// TIA Portal V19 export
DATA_BLOCK "ALL_PUMPS_DB"   // DB13
// stored: InstanceOfName ALL_PUMPS, InstanceOfType FB
"ALL_PUMPS"
   // VAR
   //    PUMP_FB1_CP01 { S7_SetPoint := 'True'} : "PUMP_FB1";
   //    PUMP_FB1_AG01 { S7_SetPoint := 'True'} : "PUMP_FB1";
   //    PUMP_FB1_CHS_CP01 { S7_SetPoint := 'True'} : "PUMP_FB1";
   //    PUMP_FB1_CHS_CP02 { S7_SetPoint := 'True'} : "PUMP_FB1";
   //    PUMP_FB1_CHS_CP03 { S7_SetPoint := 'True'} : "PUMP_FB1";
   //    PUMP_FB1_R2_CP01 { S7_SetPoint := 'True'} : "PUMP_FB1";
   //    PUMP_FB1_R2_AG01 { S7_SetPoint := 'True'} : "PUMP_FB1";
   //    PUMP_FB1_R3_CP01 { S7_SetPoint := 'True'} : "PUMP_FB1";
   //    PUMP_FB1_R3_AG01 { S7_SetPoint := 'True'} : "PUMP_FB1";
   //    PUMP_FB1_R4_CP01 { S7_SetPoint := 'True'} : "PUMP_FB1";
   //    PUMP_FB1_R4_AG01 { S7_SetPoint := 'True'} : "PUMP_FB1";
   //    PUMP_FB1_R5_CP01 { S7_SetPoint := 'True'} : "PUMP_FB1";
   //    PUMP_FB1_R5_AG01 { S7_SetPoint := 'True'} : "PUMP_FB1";
   //    PUMP_FB1_R6_CP01 { S7_SetPoint := 'True'} : "PUMP_FB1";
   //    PUMP_FB1_R6_AG01 { S7_SetPoint := 'True'} : "PUMP_FB1";
   //    PUMP_FB1_R7_CP01 { S7_SetPoint := 'True'} : "PUMP_FB1";
   //    PUMP_FB1_R7_AG01 { S7_SetPoint := 'True'} : "PUMP_FB1";
   //    PUMP_FB1_R8_CP01 { S7_SetPoint := 'True'} : "PUMP_FB1";
   //    PUMP_FB1_R8_AG01 { S7_SetPoint := 'True'} : "PUMP_FB1";
   //    PUMP_FB1_R9_CP01 { S7_SetPoint := 'True'} : "PUMP_FB1";
   //    PUMP_FB1_R9_AG01 { S7_SetPoint := 'True'} : "PUMP_FB1";
   //    PUMP_FB1_R10_CP01 { S7_SetPoint := 'True'} : "PUMP_FB1";
   //    PUMP_FB1_R10_AG01 { S7_SetPoint := 'True'} : "PUMP_FB1";
   //    PUMP_FB1_R11_CP01 { S7_SetPoint := 'True'} : "PUMP_FB1";
   //    PUMP_FB1_R11_AG01 { S7_SetPoint := 'True'} : "PUMP_FB1";
   //    PUMP_FB1_R12_CP01 { S7_SetPoint := 'True'} : "PUMP_FB1";
   //    PUMP_FB1_R12_AG01 { S7_SetPoint := 'True'} : "PUMP_FB1";
   //    PUMP_FB1_R13_CP01 { S7_SetPoint := 'True'} : "PUMP_FB1";
   //    PUMP_FB1_R13_AG01 { S7_SetPoint := 'True'} : "PUMP_FB1";
   //    PUMP_FB1_R14_CP01 { S7_SetPoint := 'True'} : "PUMP_FB1";
   //    PUMP_FB1_R14_AG01 { S7_SetPoint := 'True'} : "PUMP_FB1";
   //    PUMP_FB1_R15_CP01 { S7_SetPoint := 'True'} : "PUMP_FB1";
   //    PUMP_FB1_R15_AG01 { S7_SetPoint := 'True'} : "PUMP_FB1";
   //    PUMP_FB1_R16_CP01 { S7_SetPoint := 'True'} : "PUMP_FB1";
   //    PUMP_FB1_R16_AG01 { S7_SetPoint := 'True'} : "PUMP_FB1";
   //    PUMP_FB1_R17_CP01 { S7_SetPoint := 'True'} : "PUMP_FB1";
   //    PUMP_FB1_R17_AG01 { S7_SetPoint := 'True'} : "PUMP_FB1";
   //    PUMP_FB1_R18_CP01 { S7_SetPoint := 'True'} : "PUMP_FB1";
   //    PUMP_FB1_R18_AG01 { S7_SetPoint := 'True'} : "PUMP_FB1";
   //    PUMP_FB1_CS_CP01 { S7_SetPoint := 'True'} : "PUMP_FB1";
   //    PUMP_FB1_CS_CP02 { S7_SetPoint := 'True'} : "PUMP_FB1";
   //    PUMP_FB1_CS_CP03 { S7_SetPoint := 'True'} : "PUMP_FB1";
   //    PUMP_FB1_UCHS_CP01 { S7_SetPoint := 'True'} : "PUMP_FB1";
   //    PUMP_FB1_UCHS_CP02 { S7_SetPoint := 'True'} : "PUMP_FB1";
   //    PUMP_FB1_UCHS_CP03 { S7_SetPoint := 'True'} : "PUMP_FB1";
   //    PUMP_FB1_HS_CP01 { S7_SetPoint := 'True'} : "PUMP_FB1";
   //    PUMP_FB1_HS_CP02 { S7_SetPoint := 'True'} : "PUMP_FB1";
   //    PUMP_FB1_HS_CP03 { S7_SetPoint := 'True'} : "PUMP_FB1";
   //    "PUMP_FB1_A/SCRB_001_CP01" { S7_SetPoint := 'True'} : "PUMP_FB1";
   //    "PUMP_FB1_A/SCRB_001_CP02" { S7_SetPoint := 'True'} : "PUMP_FB1";
   //    "PUMP_FB1_A/SCRB_002_CP01" { S7_SetPoint := 'True'} : "PUMP_FB1";
   //    "PUMP_FB1_A/SCRB_001_BL01" { S7_SetPoint := 'True'} : "PUMP_FB1";
   //    "PUMP_FB1_A/SCRB_002_BL02" { S7_SetPoint := 'True'} : "PUMP_FB1";
   //    "PUMP_FB1_AA/VP_01_CP01" { S7_SetPoint := 'True'} : "PUMP_FB1";
   //    "PUMP_FB1_A/VP_01_CP01" { S7_SetPoint := 'True'} : "PUMP_FB1";
   // END_VAR
BEGIN
END_DATA_BLOCK
